FUNCTION_BLOCK COMPRESSOR
  VAR_INPUT
    PressLow   : BOOL;
    PressHigh  : BOOL;
    MinOffDone : BOOL;
  END_VAR
  VAR_OUTPUT
    Load : BOOL;
  END_VAR

BEGIN
Load := (Load OR (PressLow AND MinOffDone)) AND NOT PressHigh;
  //#ASSERT NOT (Load AND PressHigh) : P1
END_FUNCTION_BLOCK
